Fanuc KAREL source: kx00024.KL

PROGRAM KX00024
%STACKSIZE=65535
%PRIORITY=65535
%NOLOCKGROUP
VAR
I : INTEGER
J : INTEGER
B : BOOLEAN
F : FILE
S : STRING[80]
P : XYZWPR
-- UNRESOLVED DECLARATIONS (source type spelling not recovered)
-- CNF : TYPE_0x001C (type_u16=0x001C)
BEGIN
-- UNRESOLVED_PC line 12 opcodes [9D 22 A5] marker_code=0
-- UNRESOLVED_PC line 13 opcodes [22 A4 23] marker_code=15
END KX00024
